  F : ARRAY[0..5931] OF REAL := [2.842882, 6.817853, 6.893808, 6.8648725, 6.890191, 6.922743, 6.92636, 6.929977, 6.9516783, 6.915509, 6.890191, 6.9733796, 6.980613, 6.890191, 6.915509, 6.919126, 6.929977, 6.9408274, 6.929977, 6.9480615, 6.991464, 7.020399, 6.9480615, 7.005932, 6.9842305, 6.9986978, 6.991464, 6.9625287, 7.005932, 7.002315, 7.0131655, 6.980613, 7.0131655, 7.0095487, 7.0131655, 6.9733796, 7.0131655, 7.0384836, 7.060185, 7.0457177, 7.096354, 7.092737, 7.0529513, 7.071036, 7.0999713, 7.0638022, 7.1180553, 7.056568, 7.1289062, 7.143374, 7.1180553, 7.1252894, 7.172309, 7.1252894, 7.1614585, 7.0891204, 7.0999713, 7.146991, 7.2229457, 7.1180553, 7.157841, 7.1903934, 7.7654805, 8.412905, 9.027778, 9.707755, 10.304543, 10.250289, 10.235822, 10.250289, 10.304543, 10.279224, 10.358796, 10.297309, 10.420283, 10.4347515, 10.373264, 10.452836, 10.456452, 10.427517, 10.463686, 10.4817705, 10.503472, 10.521557, 10.546875, 10.583044, 10.579427, 10.619213, 10.6119795, 10.644531, 10.666233, 10.734954, 10.734954, 10.698785, 10.774739, 10.78559, 10.807292, 10.778357, 10.756655, 10.821759, 10.850695, 10.807292, 10.847077, 10.904948, 10.8723955, 10.876013, 10.944734, 10.944734, 11.009838, 11.006221, 11.020689, 11.064092, 11.035156, 11.08941, 11.118345, 11.172599, 11.158131, 11.158131, 11.125579, 11.161748, 11.2630205, 11.205151, 11.29919, 11.288339, 11.219618, 11.31004, 11.306423, 11.317274, 11.349827, 11.364294, 11.378761, 11.429399, 11.447483, 11.400463, 11.454717, 11.46195, 11.490886, 11.527055, 11.548756, 11.570457, 11.624711, 11.534288, 11.682581, 11.621094, 11.599392, 11.657263, 11.747685, 11.722367, 11.76577, 11.725984, 11.71875, 11.754919, 11.801939, 11.921296, 12.008101, 12.145544, 12.286603, 12.358941, 12.398726, 12.543403, 12.641059, 12.760417, 12.814671, 12.941261, 13.057002, 13.122107, 13.208912, 13.335504, 13.440393, 13.53805, 13.599537, 13.708044, 13.791233, 13.939526, 14.022714, 14.123987, 14.210793, 14.322917, 14.391638, 14.47121, 14.579717, 14.735243, 14.728009, 14.919704, 14.999276, 15.140336, 15.223524, 15.332031, 15.4296875, 15.530961, 15.625, 15.675636, 15.838397, 15.878182, 15.921586, 16.084347, 16.24349, 16.323061, 16.44242, 16.540075, 16.543692, 16.731771, 16.818577, 16.171152, 15.386285, 14.47121, 13.729745, 12.999132, 12.890625, 12.879774, 12.97743, 12.959346, 12.959346, 13.006366, 12.999132, 13.035301, 13.006366, 13.057002, 13.075087, 13.132957, 13.132957, 13.190827, 13.198061, 13.154658, 13.266783, 13.23423, 13.28125, 13.295717, 13.299335, 13.302952, 13.317419, 13.382524, 13.349971, 13.404224, 13.483796, 13.38614, 13.505498, 13.48018, 13.530816, 13.530816, 13.581452, 13.588686, 13.6067705, 13.632089, 13.635706, 13.661024, 13.726129, 13.711661, 13.722511, 13.726129, 13.776765, 13.740596, 13.838252, 13.831018, 13.838252, 13.906974, 13.935908, 13.932292, 13.939526, 13.986546, 13.964844, 13.993779, 14.1276045, 14.019097, 14.134838, 14.134838, 14.12037, 14.138454, 14.1276045, 14.189092, 14.254195, 14.210793, 14.210793, 14.2578125, 14.290364, 14.290364, 14.348235, 14.326533, 14.395255, 14.431423, 14.420573, 14.413339, 14.478443, 14.521846, 14.507379, 14.576099, 14.514612, 14.572483, 14.58695, 14.561632, 14.699074, 14.662905, 14.69184, 14.742476, 14.767796, 14.800347, 14.78588, 14.850984, 14.803964, 16.030092, 18.514902, 21.050346, 23.488136, 25.99103, 28.47584, 30.9932, 33.449074, 35.92303, 38.465714, 40.93967, 40.990307, 37.807438, 35.337093, 32.7908, 30.35301, 27.846498, 25.343605, 22.887732, 20.330584, 17.896412, 15.379051, 13.136574, 13.111256, 13.049768, 13.111256, 13.049768, 13.0027485, 12.973814, 12.97743, 12.86169, 12.934028, 12.890625, 12.876158, 12.876158, 12.814671, 12.839989, 12.785735, 12.774884, 12.706163, 12.760417, 12.706163, 12.666377, 12.6953125, 12.644676, 12.622974, 12.597656, 12.554254, 12.590423, 12.528935, 12.503617, 12.532552, 12.510851, 12.413195, 12.420428, 12.398726, 12.402344, 12.337239, 12.351707, 12.333623, 12.261285, 12.239583, 12.257668, 12.207031, 12.203414, 12.185329, 12.163629, 12.192564, 12.141927, 12.131077, 12.047888, 12.09129, 12.040654, 12.037037, 11.982783, 12.015336, 11.961082, 11.935764, 11.92853, 11.91768, 11.856193, 11.888744, 11.867043, 11.794704, 11.801939, 11.805555, 11.762153, 11.71875, 11.700665, 11.67173, 11.697048, 11.617476, 11.584925, 11.635561, 11.599392, 11.570457, 11.555989, 11.545139, 11.516204, 11.476418, 11.498119, 11.469184, 11.46195, 11.407697, 11.342592, 11.443866, 11.349827, 11.328125, 11.281105, 11.230469, 11.306423, 11.223235, 11.201533, 11.226851, 11.129195, 11.082176, 11.111111, 11.121962, 11.078559, 11.0496235, 11.082176, 11.006221, 11.103877, 11.038774, 10.99537, 10.933883, 10.966435, 10.915798, 10.89048, 10.854311, 10.923033, 10.814526, 10.8723955, 10.767506, 10.807292, 10.796441, 10.756655, 10.713252, 10.724103, 10.655382, 10.673467, 10.6119795, 10.666233, 10.626447, 10.554109, 10.543258, 10.507089, 10.525173, 10.489005, 10.56496, 10.507089, 10.478154, 10.420283, 10.398582, 10.398582, 10.362413, 10.369647, 10.311776, 10.347945, 10.282842, 10.297309, 10.206886, 10.275608, 10.224971, 10.243055, 10.206886, 10.127315, 10.159867, 10.134548, 10.116464, 10.123698, 10.05136, 10.127315, 10.047743, 10.040509, 10.007957, 10.018807, 10.015191, 9.888599, 9.975405, 9.910301, 9.942853, 9.895833, 9.942853, 9.859664, 9.809028, 9.812645, 9.827112, 9.758391, 9.751158, 9.769242, 9.711371, 9.689671, 9.664351, 9.686053, 9.595631, 9.617332, 9.58478, 9.57393, 9.624566, 9.5703125, 9.505208, 9.4871235, 9.490741, 9.47989, 9.469039, 9.436487, 9.393085, 9.393085, 9.385851, 9.367766, 9.324364, 9.32798, 9.313513, 9.277344, 9.288195, 9.266493, 9.255642, 9.201389, 9.201389, 9.197772, 9.215857, 9.150752, 9.150752, 9.16522, 9.161603, 9.100116, 9.085649, 8.995226, 9.016927, 9.020544, 8.984375, 8.991609, 8.96629, 8.937355, 8.95544, 8.904803, 8.89757, 8.868634, 8.901186, 8.810764, 8.79268, 8.785445, 8.832465, 8.807147, 8.709491, 8.7058735, 8.723958, 8.69864, 8.676939, 8.687789, 8.637153, 8.586516, 8.669704, 8.65162, 8.311632, 7.671441, 7.060185, 6.4127603, 5.754485, 5.5266204, 5.519387, 5.541088, 5.5266204, 5.5483217, 5.46875, 5.4904513, 5.5013022, 5.4868345, 5.494068, 5.4253473, 5.4217305, 5.479601, 5.4868345, 5.396412, 5.4253473, 5.4361978, 5.428964, 5.465133, 5.4217305, 5.432581, 5.4361978, 5.443432, 5.3855615, 5.4217305, 5.4253473, 5.432581, 5.432581, 5.3855615, 5.360243, 5.4000287, 5.3493924, 5.3385415, 5.3385415, 5.331308, 5.342159, 5.342159, 5.4108796, 5.3132234, 5.360243, 5.2987556, 5.327691, 5.3023725, 5.3023725, 5.31684, 5.31684, 5.367477, 5.280671, 5.31684, 5.2842884, 5.291522, 5.255353, 5.331308, 5.2408853, 5.3132234, 5.2842884, 5.230035, 5.2842884, 5.2336516, 5.2336516, -0.014467592, 5.295139, 7.096354, 7.0493345, 7.0782695, 7.060185, 7.0240164, 7.0999713, 7.1180553, 7.0891204, 7.060185, 7.103588, 7.13614, 7.0855036, 7.1289062, 7.1252894, 7.071036, 7.1216726, 7.1903934, 7.107205, 7.1903934, 7.146991, 7.1289062, 7.146991, 7.18316, 7.1867766, 7.1650753, 7.1903934, 7.1976275, 7.18316, 7.168692, 7.2265625, 7.18316, 7.1903934, 7.212095, 7.219329, 7.208478, 7.2229457, 7.2301793, 7.1976275, 7.2554975, 7.244647, 7.2663484, 7.269965, 7.295284, 7.2229457, 7.3350697, 7.2916665, 7.284433, 7.284433, 7.2229457, 7.306134, 7.2989006, 7.280816, 7.8993053, 8.622685, 9.186921, 9.874132, 10.438368, 10.36603, 10.380498, 10.409432, 10.441985, 10.536024, 10.550492, 10.521557, 10.521557, 10.521557, 10.597511, 10.525173, 10.630064, 10.651765, 10.640914, 10.666233, 10.698785, 10.753038, 10.78559, 10.6589985, 10.789207, 10.753038, 10.814526, 10.796441, 10.810908, 10.876013, 10.865162, 10.912182, 10.908565, 10.980903, 10.912182, 10.919415, 10.98452, 10.941117, 11.017072, 11.053241, 11.031539, 11.129195, 11.107494, 11.13643, 11.121962, 11.187066, 11.201533, 11.2160015, 11.219618, 11.288339, 11.295573, 11.244936, 11.266638, 11.338976, 11.364294, 11.302807, 11.378761, 11.407697, 11.396846, 11.433015, 11.454717, 11.480035, 11.476418, 11.501736, 11.51982, 11.505353, 11.548756, 11.588542, 11.599392, 11.6066265, 11.631945, 11.610243, 11.733217, 11.71875, 11.736835, 11.700665, 11.773004, 11.834491, 11.8308735, 11.812789, 11.812789, 11.848958, 11.877893, 11.979167, 12.076823, 12.152778, 12.225116, 12.340857, 12.3878765, 12.525318, 12.641059, 12.7568, 12.894242, 12.984664, 13.0027485, 13.161892, 13.2161455, 13.3933735, 13.454861, 13.556134, 13.70081, 13.722511, 13.859954, 13.946759, 14.084202, 14.203559, 14.344618, 14.42419, 14.568866, 14.58695, 14.702691, 14.825665, 14.963108, 15.024595, 15.1222515, 15.20544, 15.328414, 15.455006, 15.534577, 15.664786, 15.769676, 15.842014, 15.983073, 16.073496, 16.210938, 16.257957, 16.37008, 16.540075, 16.597946, 16.66305, 16.847511, 16.901766, 17.035591, 17.15133, 16.88368, 15.99754, 15.133101, 14.283131, 13.415075, 12.999132, 13.053386, 13.089555, 13.118489, 13.183594, 13.125724, 13.187211, 13.165509, 13.241464, 13.208912, 13.299335, 13.313802, 13.270399, 13.299335, 13.400608, 13.364439, 13.375289, 13.43316, 13.447627, 13.451244, 13.487413, 13.494647, 13.566985, 13.516349, 13.53805, 13.610388, 13.588686, 13.661024, 13.570601, 13.751447, 13.722511, 13.7839985, 13.744213, 13.773149, 13.773149, 13.831018, 13.794849, 13.823785, 13.917824, 13.91059, 13.841869, 14.001013, 13.928675, 13.961226, 13.986546, 14.066117, 14.01548, 14.026331, 14.12037, 14.055266, 14.149305, 14.10952, 14.1746235, 14.185474, 14.26143, 14.286748, 14.27228, 14.283131, 14.337384, 14.337384, 14.398871, 14.373553, 14.416956, 14.391638, 14.496528, 14.492911, 14.492911, 14.536314, 14.550781, 14.5652485, 14.579717, 14.623119, 14.64482, 14.623119, 14.637587, 14.684607, 14.717158, 14.782263, 14.746094, 14.728009, 14.829283, 14.89077, 14.898004, 14.916088, 14.934173, 14.934173, 14.992043, 14.999276, 15.006511, 15.049913, 15.107783, 15.118634, 15.158421, 15.143952, 15.162037, 15.198206, 15.165654, 15.219908, 15.295862, 15.259693, 15.248842, 15.350116, 15.382668, 15.389901, 15.4296875, 15.400752, 15.462239, 15.47309, 15.487557, 15.563513, 17.353878, 19.889322, 22.30541, 24.833622, 27.34375, 29.78154, 32.320602, 34.776474, 37.30107, 39.803963, 42.332176, 42.306858, 38.964844, 36.433014, 33.995224, 31.488716, 29.003906, 26.450377, 24.005354, 21.538628, 18.995949, 16.53284, 14.029948, 13.237847, 13.201678, 13.183594, 13.154658, 13.154658, 13.147425, 13.132957, 13.078704, 13.042535, 13.035301, 13.006366, 13.035301, 12.973814, 12.966579, 12.854456, 12.86169, 12.850839, 12.821904, 12.792969, 12.796586, 12.771267, 12.771267, 12.771267, 12.65191, 12.630208, 12.673611, 12.662761, 12.608507, 12.637443, 12.550636, 12.554254, 12.568721, 12.474682, 12.528935, 12.39511, 12.39511, 12.3878765, 12.402344, 12.3878765, 12.311921, 12.264901, 12.282986, 12.286603, 12.246818, 12.275752, 12.217882, 12.160011, 12.170862, 12.160011, 12.145544, 12.094908, 12.062355, 12.004485, 12.029803, 11.990017, 12.000868, 11.946614, 11.932147, 11.888744, 11.859809, 11.899595, 11.874276, 11.812789, 11.841724, 11.841724, 11.769386, 11.780237, 11.762153, 11.675347, 11.642796, 11.668114, 11.67173, 11.610243, 11.581307, 11.584925, 11.537905, 11.534288, 11.555989, 11.498119, 11.411314, 11.422164, 11.436632, 11.389612, 11.34621, 11.349827, 11.378761, 11.281105, 11.302807, 11.226851, 11.252171, 11.226851, 11.201533, 11.121962, 11.165364, 11.150897, 11.114728, 11.067708, 11.056858, 11.071325, 11.024305, 11.017072, 10.970052, 10.955585, 10.959202, 10.948351, 10.883246, 10.912182, 10.865162, 10.901331, 10.796441, 10.760272, 10.763889, 10.73857, 10.720486, 10.828993, 10.73857, 10.622829, 10.677083, 10.6119795, 10.630064, 10.590278, 10.568577, 10.51794, 10.557726, 10.51794, 10.503472, 10.463686, 10.4347515, 10.449219, 10.420283, 10.380498, 10.445601, 10.304543, 10.373264, 10.286458, 10.2683735, 10.304543, 10.246673, 10.188802, 10.264757, 10.174335, 10.152633, 10.159867, 10.120081, 10.138165, 10.09838, 10.120081, 10.083912, 10.000724, 10.047743, 9.993489, 10.018807, 9.971788, 9.950087, 9.881366, 9.89945, 9.892217, 9.856048, 9.863281, 9.856048, 9.837963, 9.758391, 9.765625, 9.78371, 9.751158, 9.704138, 9.696904, 9.635417, 9.660735, 9.642651, 9.617332, 9.610099, 9.548611, 9.552228, 9.523293, 9.497974, 9.458189, 9.490741, 9.505208, 9.472656, 9.443721, 9.411169, 9.458189, 9.403935, 9.364149, 9.335214, 9.324364, 9.320746, 9.3098955, 9.237557, 9.244792, 9.201389, 9.186921, 9.212239, 9.201389, 9.132668, 9.074798, 9.060329, 9.085649, 9.035011, 9.045862, 9.060329, 8.980758, 9.00246, 8.915654, 8.904803, 8.930121, 8.861401, 8.854167, 8.839699, 8.785445, 8.828849, 8.832465, 8.774595, 8.807147, 8.691406, 8.716724, 8.687789, 8.756511, 8.666088, 8.633536, 8.622685, 8.582899, 8.553964, 8.553964, 8.557581, 8.521412, 8.525029, 8.517796, 8.496094, 8.463542, 8.420139, 8.423756, 8.39482, 8.478009, 8.391204, 8.402055, 8.340568, 8.275463, 8.293548, 8.3152485, 8.224827, 8.297164, 8.279079, 8.087384, 7.4363427, 6.7382812, 6.14511, 5.439815, 5.1576967, 5.10706, 5.0708914, 5.114294, 5.0600405, 5.1359954, 5.078125, 5.078125, 5.1215277, 5.0962095, 5.0311055, 5.0998263, 5.0455728, 5.016638, 5.0347223, 5.0311055, 5.04919, 5.013021, 5.038339, 5.038339, 5.00217, 5.027488, 4.976852, 5.00217, 5.013021, 4.9949365, 4.969618, 4.976852, 5.005787, 4.973235, 5.016638, 5.038339, 4.9949365, 4.973235, 5.013021, 4.9913197, 4.9081306, 4.9225984, 4.9334493, 4.900897, 4.864728, 4.864728, 4.9225984, 4.890046, 4.9081306, 4.8791957, 4.9153647, 4.9479165, 4.904514, 4.868345, 4.8864293, 4.8864293, 1.7216436, 2.311198, 3.0381944, 3.656684, 3.9243345, 3.8881655, 3.8809316, 3.942419, 3.9243345, 3.982205, 3.938802, 4.0256076, 3.9858217, 4.0364585, 4.0039062, 4.0364585, 4.0039062, 4.0364585, 4.0690103, 4.1377316, 4.079861, 4.0690103, 4.1341147, 4.1413484, 4.123264, 4.170284, 4.1377316, 4.1666665, 4.1304975, 4.195602, 4.181134, 4.184751, 4.260706, 4.231771, 4.2498555, 4.3113427, 4.3113427, 4.336661, 4.3185763, 4.369213, 4.3547454, 4.3402777, 4.3764467, 4.405382, 4.3909144, 4.405382, 4.448785, 4.408999, 4.4270835, 4.398148, 4.5319734, 4.5319734, 4.5572915, 4.47772, 4.5211225, 4.546441, 4.5247397, 4.5175056, 4.6006947, 4.578993, 4.571759, 4.6043115, 4.622396, 4.662182, 4.662182, 4.7200522, 4.6694155, 4.7055845, 4.763455, 4.723669, 4.7851562, 4.7417536, 4.7453704, 4.748987, 4.788773, 4.796007, 4.788773, 4.8791957, 4.835793, 4.89728, 4.8466434, 4.926215, 4.9225984, 4.8791957, 4.9153647, 4.9189816, 4.9949365, 4.9804688, 5.0094037, 4.9985533, 5.04919, 5.1576967, 5.295139, 5.403646, 5.4470487, 5.530237, 5.6278934, 5.7689524, 5.8774595, 5.9461803, 6.000434, 6.1197915, 6.1957464, 6.311487, 6.4055266, 6.4778647, 6.5827546, 6.651476, 6.752749, 6.893808, 6.9372106, 7.0457177, 7.1506076, 7.1940103, 7.316985, 7.4363427, 7.5665507, 7.5846353, 7.700376, 7.8305845, 7.8993053, 7.96441, 8.076533, 8.105469, 8.300781, 8.369502, 8.4816265, 8.532263, 8.680555, 8.7890625, 8.886719, 8.95544, 9.0494795, 9.168837, 9.248408, 9.313513, 9.469039, 9.465423, 9.6535015, 9.725839, 9.331597, 8.5286455, 7.7256947, 6.929977, 6.0800056, 5.7689524, 5.797888, 5.758102, 5.855758, 5.848524, 5.8412905, 5.83044, 5.8449073, 5.895544, 5.9534144, 5.8810763, 5.9497976, 5.9534144, 5.910012, 5.9932003, 5.9787326, 6.032986, 5.9823494, 6.0583043, 6.047454, 6.061921, 6.047454, 6.1270256, 6.0872397, 6.1306424, 6.174045, 6.1197915, 6.1306424, 6.2319155, 6.188513, 6.2029805, 6.2174478, 6.213831, 6.2355323, 6.25, 6.3440394, 6.2970195, 6.2644677, 6.358507, 6.289786, 6.3331885, 6.3187213, 6.438079, 6.3729744, 6.3729744, 6.427228, 6.4091434, 6.4453125, 6.4561634, 6.492332, 6.4850984, 6.575521, 6.514034, 6.5610533, 6.5574365, 6.5574365, 6.6840277, 6.6225405, 6.640625, 6.61169, 6.741898, 6.6948786, 6.676794, 6.7238135, 6.6731772, 6.792535, 6.7274303, 6.7853007, 6.7599826, 6.778067, 6.778067, 6.7744503, 6.8467884, 6.890191, 6.9372106, 6.850405, 6.922743, 6.9516783, 6.9335938, 6.9480615, 6.9625287, 6.980613, 6.9842305, 7.0095487, 7.027633, 7.103588, 7.0638022, 7.0746527, 7.1144385, 7.13614, 7.143374, 7.8197336, 10.300926, 12.771267, 15.295862, 17.798756, 20.283566, 22.793692, 25.296585, 27.734375, 30.197483, 32.736546, 35.232204, 37.702545, 40.227142, 40.165653, 37.08044, 34.599247, 32.08912, 29.564526, 27.155672, 24.631077, 22.128183, 19.56742, 17.126013, 14.626736, 12.163629, 9.642651, 7.1289062, 5.4108796, 5.4144964, 5.36386, 5.353009, 5.3891783, 5.3023725, 5.287905, 5.287905, 5.3240743, 5.2336516, 5.2372684, 5.280671, 5.219184, 5.219184, 5.1359954, 5.219184, 5.179398, 5.143229, 5.143229, 5.1685476, 5.074508, 5.0925927, 5.0455728, 5.0962095, 5.027488, 4.9551506, 5.0347223, 5.0094037, 5.027488, 4.9949365, 4.9804688, 4.926215, 4.9117475, 4.962384, 4.89728, 4.875579, 4.890046, 4.8466434, 4.7743053, 4.79239, 4.8213253, 4.8177085, 4.83941, 4.796007, 4.727286, 4.716435, 4.6802664, 4.7019677, 4.6875, 4.6694155, 4.647714, 4.626013, 4.651331, 4.586227, 4.636863, 4.626013, 4.539207, 4.499421, 4.560909, 4.5428243, 4.53559, 4.5319734, 4.4560184, 4.474103, 4.474103, 4.448785, 4.5211225, 4.4632525, 4.4162326, 4.3836803, 4.336661, 4.3511286, 4.296875, 4.3185763, 4.3511286, 4.3149595, 4.3041086, 4.347512, 4.2643228, 4.271557, 4.260706, 4.235388, 4.3041086, 4.1739006, 4.188368, 4.195602, 4.159433, 4.1521993, 4.119647, 4.119647, 4.108796, 4.1015625, 4.05816, 4.123264, 4.0726275, 4.083478, 3.9605036, 4.0039062, 4.007523, 4.0256076, 3.9858217, 3.8990161, 3.9568865, 3.9171007, 3.9641204, 3.9207175, 3.9026332, 3.8773148, 3.8447628, 3.8483796, 3.8447628, 3.8266783, 3.830295, 3.804977, 3.7760417, 3.7507234, 3.7000868, 3.7543402, 3.7181714, 3.7000868, 3.69647, 3.685619, 3.6892362, 3.725405, 3.6639178, 3.6385996, 3.5879629, 3.6385996, 3.5807292, 3.59158, 3.5264757, 3.5083911, 3.5228589, 3.5300925, 3.4975405, 3.5011575, 3.4324362, 3.4252026, 3.5011575, 3.4324362, 3.410735, 3.4360533, 3.3962674, 3.374566, 3.370949, 3.3673322, 3.3528645, 3.3166957, 3.378183, 3.302228, 3.2841434, 3.294994, 3.233507, 3.2732928, 3.2045717, 3.226273, 3.1864872, 3.2045717, 3.2118056, 3.1394675, 3.157552, 3.161169, 3.1358507, 3.1286168, 3.1286168, 3.0454283, 3.0635128, 3.0996816, 3.0454283, 3.049045, 3.049045, 3.023727, 3.0092592, 2.9513888, 2.9513888, 2.983941, 2.980324, 2.9296875, 2.911603, 2.8573496, 2.8645833, 2.9188368, 2.911603, 2.8175638, 2.8537326, 2.842882, 2.8320312, 2.7958622, 2.7777777, 2.8139467, 2.734375, 2.7199075, 2.7596934, 2.7162905, 2.698206, 2.7416089, 2.6945891, 2.6801214, 2.6728878, 2.6367188, 2.629485, 2.6801214, 2.6367188, 2.6150174, 2.5752316, 2.564381, 2.55353, 2.5788484, 2.5426793, 2.4920428, 2.5282118, 2.5065105, 2.5028934, 2.4775753, 2.44864, 2.4088542, 2.4233217, 2.5065105, 2.3980036, 2.445023, 2.3582175, 2.4233217, 2.3618345, 2.376302, 2.3654513, 2.2858796, 2.3184316, 2.23886, 2.3365161, 2.275029, 2.2605612, 2.1918402, 2.2280092, 1.634838, 0.9765625, 0.30020255, 3.4432871, 5.0455728, 5.0998263, 5.10706, 5.0853586, 5.1613135, 5.117911, 5.128762, 5.0925927, 5.143229, 5.0600405, 5.0708914, 5.1649303, 5.128762, 5.114294, 5.103443, 5.1576967, 5.183015, 5.117911, 5.1576967, 5.179398, 5.1649303, 5.0708914, 5.1251445, 5.215567, 5.179398, 5.2119503, 5.1721644, 5.204716, 5.150463, 5.204716, 5.179398, 5.190249, 5.1974826, 5.2445025, 5.2408853, 5.1757812, 5.251736, 5.280671, 5.2445025, 5.255353, 5.2842884, 5.2408853, 5.280671, 5.2445025, 5.2336516, 5.2987556, 5.230035, 5.2698207, 5.31684, 5.3783274, 5.3385415, 5.2987556, 5.287905, 5.3132234, 5.2770543, 5.3747106, 5.3132234, 5.4000287, 5.353009, 5.3096066, 5.6315103, 6.3368053, 6.969763, 7.60272, 8.282697, 8.427373, 8.405671, 8.445457, 8.456307, 8.423756, 8.510561, 8.539496, 8.564815, 8.496094, 8.59375, 8.600984, 8.619068, 8.557581, 8.691406, 8.669704, 8.691406, 8.738426, 8.637153, 8.763744, 8.781829, 8.796296, 8.785445, 8.80353, 8.843316, 8.854167, 8.875868, 8.843316, 8.908421, 8.937355, 8.9192705, 9.006077, 8.959057, 8.998842, 8.973524, 9.016927, 9.031395, 9.031395, 8.998842, 9.085649, 9.063947, 9.154369, 9.186921, 9.161603, 9.273726, 9.201389, 9.226707, 9.233941, 9.248408, 9.248408, 9.338831, 9.338831, 9.349682, 9.302662, 9.364149, 9.447338, 9.367766, 9.454572, 9.385851, 9.42202, 9.476274, 9.490741, 9.505208, 9.505208, 9.602864, 9.555845, 9.544994, 9.588397, 9.628182, 9.664351, 9.628182, 9.660735, 9.682436, 9.729456, 9.707755, 9.73669, 9.740307, 9.823495, 9.805411, 9.798177, 9.823495, 9.866899, 9.881366, 9.85243, 9.975405, 10.007957, 9.95732, 10.029658, 10.185185, 10.206886, 10.315393, 10.467303, 10.554109, 10.691551, 10.756655, 10.789207, 10.966435, 11.067708, 11.161748, 11.205151, 11.338976, 11.472801, 11.555989, 11.603009, 11.715133, 11.794704, 11.924913, 12.040654, 12.131077, 12.203414, 12.355324, 12.384259, 12.507234, 12.60489, 12.648293, 12.800202, 12.9557295, 13.042535, 13.078704, 13.165509, 13.32827, 13.404224, 13.527199, 13.58507, 13.726129, 13.820168, 13.968461, 13.990162, 14.134838, 14.21441, 14.279514, 14.362702, 14.532697, 14.619502, 14.7316265, 14.840133, 14.923322, 14.623119, 13.798467, 12.9557295, 12.160011, 11.382379, 11.020689, 11.053241, 11.121962, 11.107494, 11.143663, 11.121962, 11.150897, 11.14728, 11.219618, 11.190682, 11.183449, 11.223235, 11.302807, 11.295573, 11.255787, 11.364294, 11.317274, 11.375145, 11.3932295, 11.418548, 11.4402485, 11.469184, 11.436632, 11.494502, 11.494502, 11.588542, 11.555989, 11.559607, 11.603009, 11.617476, 11.617476, 11.704283, 11.693432, 11.678964, 11.715133, 11.744068, 11.773004, 11.758536, 11.816406, 11.809173, 11.848958, 11.910445, 11.950232, 11.874276, 11.932147, 11.924913, 11.968316, 11.979167, 12.004485, 12.037037, 12.000868, 12.123842, 12.105758, 12.181713, 12.141927, 12.203414, 12.13831, 12.203414, 12.239583, 12.250434, 12.2432, 12.29022, 12.326389, 12.366175, 12.362557, 12.358941, 12.3878765, 12.3878765, 12.424046, 12.405961, 12.485533, 12.528935, 12.528935, 12.528935, 12.54702, 12.554254, 12.615741, 12.619358, 12.626592, 12.662761, 12.6953125, 12.764033, 12.811053, 12.724248, 12.760417, 12.80382, 12.843605, 12.836371, 12.850839, 12.90871, 12.941261, 13.292101, 15.704572, 18.17853, 20.706741, 23.1807, 25.672743, 28.121384, 30.671297, 33.15249, 35.633682, 38.151043, 40.588833, 40.559895, 37.492767, 34.964554, 32.508682, 30.016638, 27.50651, 25.043404, 22.518808, 20.070168, 17.520254, 15.089699, 12.579572, 11.237702, 11.161748, 11.2160015, 11.114728, 11.100261, 11.121962, 11.096643, 11.085793, 11.031539, 11.024305, 11.056858, 10.951967, 11.020689, 10.944734, 10.912182, 10.901331, 10.87963, 10.8253765, 10.803675, 10.789207, 10.73857, 10.745805, 10.781974, 10.706018, 10.724103, 10.593895, 10.673467, 10.6807, 10.572193, 10.554109, 10.579427, 10.503472, 10.521557, 10.52879, 10.463686, 10.445601, 10.46007, 10.532408, 10.420283, 10.35518, 10.322627, 10.326244, 10.3515625, 10.286458, 10.250289, 10.243055, 10.228588, 10.2213545, 10.181568, 10.206886, 10.192419, 10.083912, 10.112847, 10.083912, 10.054976, 10.047743, 10.007957, 10.007957, 9.964555, 9.982639, 9.986256, 9.924768, 9.89945, 9.892217, 9.848814, 9.837963, 9.884983, 9.801794, 9.780092, 9.780092, 9.754774, 9.725839, 9.725839, 9.711371, 9.693287, 9.6535015, 9.617332, 9.628182, 9.599248, 9.566695, 9.610099, 9.57393, 9.508825, 9.4871235, 9.443721, 9.414786, 9.43287, 9.382234, 9.382234, 9.360533, 9.324364, 9.338831, 9.306279, 9.378617, 9.244792, 9.215857, 9.2628765, 9.291811, 9.186921, 9.183305, 9.190538, 9.194155, 9.147136, 9.067564, 9.035011, 9.009693, 9.103733, 8.991609, 9.009693, 9.009693, 8.991609, 9.027778, 8.933739, 8.8722515, 8.933739, 8.865017, 8.875868, 8.843316, 8.7890625, 8.843316, 8.74566, 8.713108, 8.767361, 8.7058735, 8.687789, 8.673322, 8.7058735, 8.600984, 8.597367, 8.604601, 8.600984, 8.575665, 8.532263, 8.532263, 8.521412, 8.553964, 8.5286455, 8.478009, 8.4816265, 8.470776, 8.409288, 8.351418, 8.308015, 8.362268, 8.3152485, 8.3152485, 8.297164, 8.293548, 8.213976, 8.206742, 8.199508, 8.224827, 8.192274, 8.17419, 8.18504, 8.134404, 8.101851, 8.065682, 8.080151, 8.065682, 8.065682, 8.025897, 7.9716434, 8.036748, 7.9318576, 7.939091, 7.949942, 7.913773, 7.9029226, 7.8703704, 7.884838, 7.8956885, 7.837818, 7.8052664, 7.747396, 7.7582464, 7.7256947, 7.7546296, 7.703993, 7.6931424, 7.7293115, 7.6678243, 7.6171875, 7.5882525, 7.6497397, 7.5810184, 7.573785, 7.5810184, 7.530382, 7.5520835, 7.5050635, 7.486979, 7.472512, 7.5014467, 7.396557, 7.382089, 7.458044, 7.360388, 7.3423033, 7.349537, 7.309751, 7.3025174, 7.248264, 7.306134, 7.269965, 7.2265625, 7.1903934, 7.157841, 7.2012444, 7.139757, 7.168692, 7.1108217, 7.081887, 7.0746527, 7.0999713, 7.0457177, 7.1759257, 7.027633, 7.03125, 6.9878473, 6.9733796, 7.0131655, 6.929977, 6.8757234, 6.8974247, 6.857639, 6.8467884, 6.8865743, 6.8106194, 6.7599826, 6.792535, 6.814236, 6.792535, 6.2970195, 5.6351275, 4.875579, 4.257089, 3.6639178, 3.7073207, 3.69647, 3.6385996, 3.692853, 3.685619, 3.660301, 3.6639178, 3.6385996, 3.656684, 3.7181714, 3.685619, 3.6422164, 3.6277487, 3.620515, 3.6458333, 3.6385996, 3.5951967, 3.584346, 3.6313658, 3.5988138, 3.5879629, 3.5807292, 3.5879629, 3.5554109, 3.5879629, 3.59158, 3.551794, 3.5300925, 3.6060474, 3.5554109, 3.5300925, 3.5409434, 3.5264757, 3.5047743, 3.5192418, 3.5083911, 3.5373263, 3.5626447, 3.5011575, 3.5409434, 3.4866898, 3.5662615, 3.5120082, 3.5047743, 3.5192418, 3.4903066, 3.5228589, 3.4866898, 3.4505208, 3.4722223, 3.4649885, 3.446904, 3.4577546, 3.3528645, 3.4939237, 3.4866898, 3.4179688, 3.4215856, 3.4252026, 3.378183, 1.8916377, 4.615162, 4.626013, 4.5645256, 4.6187787, 4.6187787, 4.560909, 4.662182, 4.6296296, 4.6187787, 4.615162, 4.5645256, 4.622396, 4.6079283, 4.658565, 4.683883, 4.622396, 4.6043115, 4.691117, 4.6875, 4.676649, 4.647714, 4.6440973, 4.651331, 4.691117, 4.5898438, 4.6043115, 4.6730323, 4.723669, 4.6332464, 4.6730323, 4.7019677, 4.727286, 4.698351, 4.7019677, 4.6875, 4.6802664, 4.6730323, 4.6802664, 4.716435, 4.6947336, 4.6549478, 4.727286, 4.7345195, 4.738137, 4.727286, 4.788773, 4.7815394, 4.788773, 4.7670717, 4.7706885, 4.799624, 4.738137, 4.738137, 4.8177085, 4.763455, 4.8574944, 4.7815394, 4.7670717, 4.796007, 4.803241, 4.9479165, 5.5917244, 6.2934027, 6.919126, 7.526765, 7.8956885, 7.8920717, 7.8920717, 7.939091, 7.9029226, 7.960793, 7.960793, 7.960793, 7.9788775, 7.96441, 7.9463253, 8.036748, 8.018663, 8.087384, 8.065682, 8.105469, 8.141638, 8.188658, 8.145255, 8.181423, 8.192274, 8.17419, 8.275463, 8.206742, 8.199508, 8.308015, 8.257379, 8.311632, 8.326099, 8.33695, 8.322483, 8.33695, 8.3152485, 8.412905, 8.380353, 8.344184, 8.463542, 8.412905, 8.467158, 8.459925, 8.525029, 8.496094, 8.499711, 8.568432, 8.499711, 8.575665, 8.564815, 8.619068, 8.626302, 8.684173, 8.629919, 8.684173, 8.69864, 8.662471, 8.713108, 8.716724, 8.785445, 8.774595, 8.785445, 8.7890625, 8.79268, 8.846932, 8.825232, 8.904803, 8.890336, 8.930121, 8.987992, 8.973524, 8.944589, 8.933739, 9.07118, 9.01331, 9.038629, 9.020544, 9.056713, 9.07118, 9.038629, 9.125434, 9.1182, 9.103733, 9.190538, 9.139901, 9.215857, 9.244792, 9.226707, 9.284577, 9.302662, 9.400318, 9.519676, 9.602864, 9.696904, 9.801794, 9.870515, 9.94647, 10.058594, 10.174335, 10.275608, 10.380498, 10.456452, 10.568577, 10.698785, 10.745805, 10.836226, 10.944734, 11.078559, 11.085793, 11.248553, 11.367911, 11.458333, 11.530671, 11.621094, 11.700665, 11.841724, 11.92853, 12.029803, 12.152778, 12.207031, 12.344474, 12.377026, 12.518085, 12.637443, 12.713397, 12.811053, 12.883391, 13.064236, 13.089555, 13.22338, 13.292101, 13.436776, 13.527199, 13.610388, 13.718895, 13.820168, 13.932292, 14.001013, 14.073351, 13.943142, 13.136574, 12.380642, 11.563224, 10.662616, 10.199653, 10.206886, 10.275608, 10.264757, 10.257524, 10.271991, 10.282842, 10.322627, 10.402199, 10.3515625, 10.36603, 10.423901, 10.470921, 10.489005, 10.478154, 10.536024, 10.525173, 10.521557, 10.539641, 10.568577, 10.622829, 10.604745, 10.640914, 10.63368, 10.615596, 10.6589985, 10.698785, 10.767506, 10.687934, 10.724103, 10.78559, 10.807292, 10.854311, 10.756655, 10.821759, 10.774739, 10.876013, 10.857928, 10.894097, 10.857928, 10.926649, 10.930266, 10.988136, 11.035156, 11.046007, 11.038774, 11.017072, 11.096643, 11.118345, 11.085793, 11.143663, 11.201533, 11.1943, 11.201533, 11.176215, 11.230469, 11.205151, 11.342592, 11.291956, 11.31004, 11.313658, 11.313658, 11.331742, 11.41493, 11.443866, 11.407697, 11.46195, 11.447483, 11.490886, 11.51982, 11.541522, 11.545139, 11.501736, 11.628327, 11.621094, 11.628327, 11.639178, 11.624711, 11.646412, 11.682581, 11.729601, 11.71875, 11.791088, 11.794704, 11.856193, 11.834491, 11.780237, 11.845342, 11.852575, 11.859809, 11.932147, 12.084057, 14.369936, 16.880064, 19.382957, 21.849682, 24.374277, 26.837385, 29.394531, 31.807003, 34.324364, 36.816406, 39.304832, 41.82581, 41.822193, 38.697193, 36.23047, 33.716724, 31.210215, 28.68562, 26.182726, 23.672598, 21.216724, 18.75, 16.26519, 13.75868, 11.2160015, 10.21412, 10.170717, 10.199653, 10.116464, 10.058594, 10.112847, 10.073061, 10.10923, 10.080296, 9.993489, 10.015191, 10.040509, 9.968171, 9.928386, 9.924768, 9.982639, 9.942853, 9.859664, 9.870515, 9.845197, 9.845197, 9.834346, 9.85243, 9.686053, 9.765625, 9.725839, 9.73669, 9.718605, 9.7005205, 9.671586, 9.628182, 9.613715, 9.599248, 9.508825, 9.519676, 9.508825, 9.47989, 9.530526, 9.505208, 9.4401045, 9.461805, 9.458189, 9.396702, 9.360533, 9.389467, 9.295428, 9.331597, 9.306279, 9.284577, 9.313513, 9.233941, 9.295428, 9.230324, 9.226707, 9.215857, 9.136285, 9.129051, 9.0964985, 9.1182, 9.0964985, 9.056713, 9.085649, 9.042245, 9.016927, 8.998842, 9.006077, 8.959057, 8.995226, 8.933739, 8.886719, 8.868634, 8.868634, 8.886719, 8.861401, 8.825232, 8.846932, 8.723958, 8.7890625, 8.74566, 8.716724, 8.676939, 8.64077, 8.695024, 8.65162, 8.637153, 8.648004, 8.64077, 8.615452, 8.586516, 8.568432, 8.539496, 8.539496, 8.470776, 8.532263, 8.423756, 8.430989, 8.44184, 8.365886, 8.485243, 8.344184, 8.373119, 8.304399, 8.355035, 8.3152485, 8.300781, 8.246528, 8.297164, 8.257379, 8.235677, 8.206742, 8.199508, 8.177807, 8.159722, 8.152489, 8.065682, 8.148871, 8.083767, 8.065682, 8.051215, 8.047599, 8.029514, 8.01143, 7.9824944, 7.9571757, 7.9427085, 7.921007, 7.924624, 7.888455, 7.8956885, 7.8450522, 7.816117, 7.8305845, 7.873987, 7.7944155, 7.7980323, 7.675058, 7.751013, 7.736545, 7.675058, 7.6569734, 7.7329283, 7.664207, 7.6822915, 7.624421, 7.624421, 7.599103, 7.5810184, 7.5774016, 7.533999, 7.494213, 7.548466, 7.4652777, 7.530382, 7.4905963, 7.3893228, 7.411024, 7.3676214, 7.458044, 7.411024, 7.3350697, 7.3314524, 7.313368, 7.309751, 7.3025174, 7.2663484, 7.284433, 7.2374134, 7.233796, 7.244647, 7.219329, 7.132523, 7.143374, 7.143374, 7.096354, 7.0746527, 7.1289062, 7.0638022, 7.1252894, 7.0529513, 7.0638022, 7.027633, 6.9444447, 7.0638022, 6.9769964, 6.9408274, 6.966146, 6.9625287, 6.893808, 6.9625287, 6.890191, 6.890191, 6.8721066, 6.8359375, 6.8033853, 6.7997684, 6.745515, 6.749132, 6.781684, 6.702112, 6.7853007, 6.7382812, 6.7093463, 6.6731772, 6.629774, 6.6478586, 6.589988, 6.6080728, 6.6623263, 6.604456, 6.5502024, 6.5502024, 6.528501, 6.4742475, 6.503183, 6.463397, 6.4561634, 6.430845, 6.4199944, 6.4344616, 6.488715, 6.3946757, 6.391059, 6.311487, 6.351273, 6.3187213, 6.351273, 6.3078704, 6.275318, 6.2825522, 6.300637, 6.2355323, 6.25, 6.1957464, 5.5157695, 4.9189816, 4.235388, 3.6639178, 3.1394675, 3.125, 3.125, 3.092448, 3.0996816, 3.1141493, 3.1141493, 3.1213832, 3.0743635, 3.1032987, 3.092448, 3.1141493, 3.0996816, 3.1286168, 3.0381944, 3.1177661, 3.1539352, 3.0996816, 3.0635128, 3.0779803, 3.1032987, 3.0743635, 3.0309606, 3.02011, 3.0960648, 3.0635128, 3.092448, 3.0418112, 3.0526621, 3.0454283, 3.0707464, 3.0309606, 3.0345776, 3.0273438, 3.0128763, 3.0671296, 3.0020254, 3.0418112, 3.0526621, 2.9911747, 2.983941, 3.016493, 3.0598958, 3.0598958, 3.0418112, 2.9947917, 2.9911747, 3.0020254, 3.023727, 2.9911747, 2.9947917, 3.0056424, 2.9947917, 2.9767072, 2.947772, 2.9694734, 2.9694734, 2.947772, 2.9730902, 3.023727, 0.003616898, 3.8917825, 7.8667536, 10.387732, 10.405816, 10.4347515, 10.358796, 10.4347515, 10.423901, 10.423901, 10.405816, 10.391349, 10.441985, 10.423901, 10.427517, 10.445601, 10.46007, 10.463686, 10.507089, 10.4347515, 10.427517, 10.496239, 10.456452, 10.478154, 10.463686, 10.496239, 10.496239, 10.4817705, 10.416667, 10.499855, 10.51794, 10.525173, 10.532408, 10.489005, 10.507089, 10.532408, 10.496239, 10.52879, 10.590278, 10.507089, 10.550492, 10.543258, 10.561342, 10.604745, 10.590278, 10.57581, 10.601129, 10.554109, 10.543258, 10.57581, 10.604745, 10.666233, 10.640914, 10.604745, 10.6119795, 10.622829, 10.6119795, 10.63368, 10.637298, 10.669849, 10.6589985, 10.626447, 10.6807, 10.912182, 11.490886, 12.087673, 12.807436, 13.472945, 13.718895, 13.733362, 13.75868, 13.827401, 13.834636, 13.878038, 13.8671875, 13.906974, 13.86357, 13.896123, 13.928675, 13.982928, 13.964844, 14.00463, 13.939526, 14.037182, 14.033565, 14.102286, 14.1276045, 14.080585, 14.1276045, 14.102286, 14.171007, 14.156539, 14.1746235, 14.210793, 14.221643, 14.265046, 14.239728, 14.268663, 14.279514, 14.333767, 14.297599, 14.312066, 14.355469, 14.362702, 14.406105, 14.402489, 14.409722, 14.514612, 14.48206, 14.500145, 14.510995, 14.456742, 14.525463, 14.561632, 14.63397, 14.58695, 14.615886, 14.63397, 14.688224, 14.655671, 14.670139, 14.713542, 14.709925, 14.775029, 14.782263, 14.800347, 14.811198, 14.847367, 14.9088545, 14.854601, 14.869068, 14.90162, 14.934173, 14.923322, 14.959491, 14.945024, 15.002893, 15.028212, 15.05353, 15.0390625, 15.071614, 15.060764, 15.075232, 15.143952, 15.140336, 15.165654, 15.172888, 15.194589, 15.212673, 15.237992, 15.230758, 15.274161, 15.292245, 15.259693, 15.436921, 15.47309, 15.56713, 15.704572, 15.809462, 15.925202, 15.99754, 16.040943, 16.229021, 16.29051, 16.413485, 16.45327, 16.594328, 16.735388, 16.771557, 16.945168, 16.974104, 17.086227, 17.126013, 17.256222, 17.386429, 17.520254, 17.563658, 17.690248, 17.82769, 17.914497, 17.939816, 18.051939, 18.171297, 18.254484, 18.381077, 18.525753, 18.612558, 18.663195, 18.757235, 18.898293, 18.981482, 19.089989, 19.245516, 19.288918, 19.433594, 19.560184, 19.599972, 19.62529, 19.806135, 19.896557, 19.979746, 20.120804, 20.225695, 20.330584, 20.272715, 19.480614, 18.565538, 17.856627, 17.006655, 16.485823, 16.44242, 16.550926, 16.456886, 16.540075, 16.56901, 16.554543, 16.608797, 16.597946, 16.659433, 16.71007, 16.724537, 16.735388, 16.677517, 16.728153, 16.735388, 16.861979, 16.796875, 16.83666, 16.847511, 16.854746, 16.912615, 16.876448, 16.959635, 17.006655, 16.934317, 16.988571, 16.988571, 17.01389, 17.089844, 17.158566, 17.078993, 17.158566, 17.122396, 17.205584, 17.227285, 17.24537, 17.216434, 17.238136, 17.31409, 17.30324, 17.364729, 17.346643, 17.433449, 17.4443, 17.415365, 17.386429, 17.404514, 17.45515, 17.509403, 17.534721, 17.574509, 17.574509, 17.545572, 17.603443, 17.635996, 17.668547, 17.730034, 17.733652, 17.730034, 17.766203, 17.831308, 17.798756, 17.849392, 17.824074, 17.914497, 17.892796, 17.939816, 17.943432, 18.00492, 18.019386, 18.041088, 18.055555, 18.023003, 18.091724, 18.149595, 18.124277, 18.185764, 18.214699, 18.17853, 18.2364, 18.258102, 18.27257, 18.315971, 18.315971, 18.381077, 18.359375, 18.370226, 18.471498, 18.48235, 18.467882, 18.4932, 20.554832, 23.021557, 25.56062, 27.987558, 30.50492, 33.062065, 35.467304, 37.94126, 40.46224, 40.505642, 36.4511, 32.461662, 29.644096, 27.083334, 24.660011, 22.063078, 19.632523, 17.111546, 14.594184, 12.149161, 9.8307295, 9.42202, 9.497974, 9.436487, 9.360533, 9.367766, 9.302662, 9.299046, 9.2628765, 9.324364, 9.230324, 9.2628765, 9.201389, 9.248408, 9.161603, 9.139901, 9.129051, 9.129051, 9.053096, 9.082031, 9.038629, 9.01331, 8.987992, 8.95544, 8.940972, 8.940972, 8.9192705, 8.904803, 8.901186, 8.915654, 8.828849, 8.832465, 8.810764, 8.79268, 8.738426, 8.752893, 8.749276, 8.65162, 8.669704, 8.65162, 8.626302, 8.586516, 8.633536, 8.575665, 8.586516, 8.5286455, 8.470776, 8.434607, 8.430989, 8.478009, 8.409288, 8.365886, 8.33695, 8.409288, 8.333333, 8.344184, 8.347801, 8.318866, 8.322483, 8.308015, 8.192274, 8.250145, 8.206742, 8.192274, 8.163339, 8.058449, 8.105469, 8.112702, 8.047599, 8.029514, 8.080151, 8.015046, 8.0078125, 7.91739, 8.015046, 7.9318576, 7.8956885, 7.8993053, 7.8667536, 7.928241, 7.837818, 7.9065394, 7.7690973, 7.837818, 7.7907987, 7.7437787, 7.7437787, 7.740162, 7.664207, 7.7220774, 7.635272, 7.609954, 7.6063366, 7.6280384, 7.573785, 7.5665507, 7.5159144, 7.5014467, 7.4544272, 7.5050635, 7.4761286, 7.425492, 7.4399595, 7.39294, 7.411024, 7.385706, 7.3350697, 7.3350697, 7.3386865, 7.273582, 7.284433, 7.2663484, 7.2301793, 7.2157116, 7.1976275, 7.157841, 7.1940103, 7.1867766, 7.139757, 7.1144385, 7.096354, 7.081887, 7.0638022, 7.034867, 7.060185, 6.9842305, 6.854022, 6.980613, 6.9408274, 6.929977, 6.904659, 6.9118924, 6.82147, 6.828704, 6.817853, 6.778067, 6.7961516, 6.7310476, 6.7853007, 6.778067, 6.702112, 6.665943, 6.680411, 6.629774, 6.579138, 6.6225405, 6.6550927, 6.5863714, 6.640625, 6.5502024, 6.5610533, 6.514034, 6.467014, 6.4814816, 6.4959493, 6.45978, 6.430845, 6.391059, 6.35489, 6.391059, 6.358507, 6.362124, 6.35489, 6.35489, 6.289786, 6.25, 6.1921296, 6.239149, 6.221065, 6.1921296, 6.1704283, 6.1306424, 6.1631947, 6.1306424, 6.112558, 6.141493, 6.069155, 6.0149016, 6.0257525, 6.0149016, 5.9136286, 5.996817, 5.964265, 5.920862, 5.964265, 5.862992, 5.9136286, 5.870226, 5.8521414, 5.834057, 5.8521414, 5.808738, 5.794271, 5.797888, 5.7725697, 5.7038484, 5.721933, 5.6893806, 5.6532116, 5.721933, 5.67853, 5.6387444, 5.6025753, 5.5664062, 5.5627894, 5.5013022, 5.5483217, 5.4832177, 5.497685, 5.497685, 5.4615164, 5.479601, 5.443432, 5.4361978, 5.392795, 5.3819447, 5.3710938, 5.327691, 5.255353, 5.3132234, 5.2408853, 5.186632, 5.291522, 5.2481194, 5.2372684, 5.2372684, 5.2010994, 5.1974826, 5.1721644, 5.1757812, 5.15408, 5.15408, 5.0962095, 4.9153647, 4.2426214, 3.584346, 2.983941, 2.3039641, 2.0182292, 1.9675926, 1.9929109, 2.0073786, 2.0146122, 1.9748263, 1.9856771, 1.9024885, 1.9712095, 1.8952546, 1.9675926, 1.9748263, 1.9241898, 1.9567419, 1.9458913, 1.9422743, 1.9748263, 1.8735533, 1.9024885, 1.9205729, 1.9241898, 1.9133391, 1.880787, 1.9350405, 1.9567419, 1.8590857, 1.9024885, 1.8880209, 1.8373842, 1.8590857, 1.884404, 1.8699363, 1.8265336, 1.8229166, 1.812066, 1.8554688, 1.8554688, 1.848235, 1.848235, 1.8590857, 1.8265336, 1.775897, 1.8446181, 1.8192998, 1.7903646, 1.8301505, 1.8554688, 1.7903646, 1.739728, 1.8012153, 1.7614294, 1.808449, 1.775897, 1.7469618, 1.7505788, 1.8012153, 1.7650462, 1.7722801, 1.7433449, 1.775897, 2.665654, 6.741898, 6.904659, 6.915509, 6.980613, 6.9625287, 6.8612556, 6.958912, 6.904659, 6.8721066, 6.922743, 6.9372106, 6.929977, 6.955295, 6.9372106, 6.87934, 6.904659, 6.9625287, 6.966146, 6.922743, 6.9625287, 6.92636, 6.958912, 7.0167823, 6.966146, 7.071036, 6.958912, 7.002315, 6.969763, 6.9769964, 6.9842305, 7.0131655, 7.005932, 7.020399, 7.0999713, 7.067419, 7.0384836, 7.0240164, 7.0167823, 7.0384836, 7.060185, 7.0782695, 7.0999713, 7.071036, 7.139757, 7.0891204, 7.0384836, 7.081887, 7.103588, 7.1614585, 7.1216726, 7.1180553, 7.092737, 7.157841, 7.1542244, 7.13614, 7.1614585, 7.107205, 7.18316, 7.146991, 7.2012444, 7.1940103, 7.1903934, 7.107205, 7.2012444, 7.1506076, 7.18316, 7.179543, 7.1903934, 7.1903934, 7.233796, 7.1940103, 7.2012444, 7.2157116, 7.2012444, 7.204861, 7.2518806, 7.269965, 7.2157116, 7.2229457, 7.244647, 7.2916665, 7.24103, 7.2916665, 7.295284, 7.295284, 7.2627316, 7.2518806, 7.3025174, 7.3025174, 7.306134, 7.24103, 7.2916665, 7.313368, 7.418258, 7.3242188, 7.4001737, 7.284433, 7.349537, 7.3386865, 7.3278356, 7.3784723, 7.313368, 7.425492, 7.3748555, 7.3784723, 7.4074073, 7.3640046, 7.418258, 7.4291086, 7.3640046, 7.4001737, 7.421875, 7.3784723, 7.4399595, 7.45081, 7.4037905, 7.4291086, 7.4001737, 7.4652777, 7.4761286, 7.458044, 7.472512, 7.4761286, 7.5014467, 7.4797454, 7.5014467, 7.4363427, 7.4761286, 7.5014467, 7.5159144, 7.5195312, 7.486979, 7.526765, 7.5448494, 7.533999, 7.5448494, 7.570168, 7.5520835, 7.548466, 7.548466, 7.5557003, 7.562934, 7.559317, 7.5810184, 7.60272, 7.526765, 7.5557003, 7.595486, 7.5882525, 7.6533566, 7.6171875, 7.6171875, 7.6425056, 7.6497397, 7.6280384, 7.6497397, 7.6533566, 7.6822915, 7.6533566, 7.703993, 7.696759, 7.70761, 7.6822915, 7.675058, 7.696759, 7.7582464, 7.7220774, 7.6931424, 7.7220774, 7.7329283, 7.7582464, 7.7546296, 7.7220774, 7.7293115, 7.7582464, 7.7293115, 7.761863, 7.7437787, 7.7256947, 7.7582464, 7.7980323, 7.7944155, 7.772714, 7.8595195, 7.837818, 7.8305845, 7.7980323, 7.877604, 7.837818, 7.8812213, 7.9354744, 7.877604, 7.921007, 7.8812213, 7.9029226, 7.949942, 7.8956885, 7.888455, 7.921007, 7.873987, 7.913773, 7.8920717, 7.924624, 7.939091, 7.9354744, 7.939091, 7.9571757, 7.949942, 7.9716434, 7.96441, 7.9824944, 8.02228, 7.993345, 8.047599, 7.989728, 7.986111, 8.058449, 8.015046, 8.087384, 7.9788775, 8.029514, 8.029514, 8.015046, 8.051215, 8.000579, 8.065682, 8.036748, 8.101851, 8.130787, 8.0910015, 8.098235, 8.087384, 8.109086, 8.134404, 8.072917, 8.130787, 8.152489, 8.159722, 8.159722, 8.141638, 8.181423, 8.152489, 8.134404, 8.18504, 8.156105, 8.253761, 8.210359, 8.206742, 8.286314, 8.250145, 8.264612, 8.239294, 8.250145, 8.264612, 8.257379, 8.28993, 8.28993, 8.260995, 8.2682295, 8.326099, 8.3152485, 8.39482, 8.322483, 8.293548, 8.297164, 8.308015, 8.344184, 8.369502, 8.333333, 8.412905, 8.39482, 8.402055, 8.402055, 8.467158, 8.412905, 8.412905, 8.420139, 8.423756, 8.463542, 8.456307, 8.449074, 8.391204, 8.53588, 8.459925, 8.496094, 8.48886, 8.430989, 8.532263, 8.510561, 8.474392, 8.53588, 8.525029, 8.582899, 8.525029, 8.532263, 8.550347, 8.770978, 11.060474, 13.581452, 16.04456, 18.518518, 21.097366, 23.53154, 26.016348, 28.468605, 31.011284, 33.52141, 35.991753, 38.43316, 40.91797, 40.99754, 37.7785, 35.380497, 32.816116, 30.349392, 27.81033, 25.347221, 22.858797, 20.413773, 17.86386, 15.350116, 12.91956, 10.376881, 7.96441, 6.8250866, 6.8612556, 6.8106194, 6.8359375, 6.8395543, 6.8106194, 6.792535, 6.8106194, 6.7744503, 6.7853007, 6.792535, 6.756366, 6.7744503, 6.7274303, 6.7382812, 6.756366, 6.767216, 6.749132, 6.6876445, 6.7635994, 6.7708335, 6.7093463, 6.702112, 6.741898, 6.691262, 6.640625, 6.6948786, 6.6333914, 6.640625, 6.604456, 6.651476, 6.640625, 6.6478586, 6.600839, 6.5936055, 6.6080728, 6.5863714, 6.5863714, 6.6080728, 6.6225405, 6.6189237, 6.579138, 6.615307, 6.6080728, 6.5610533, 6.6225405, 6.528501, 6.5502024, 6.524884, 6.492332, 6.528501, 6.5104165, 6.532118, 6.4453125, 6.488715, 6.4489293, 6.488715, 6.4778647, 6.4706306, 6.463397, 6.40191, 6.4344616, 6.4453125, 6.4416957, 6.4489293, 6.387442, 6.4091434, 6.423611, 6.40191, 6.427228, 6.427228, 6.3946757, 6.376591, 6.45978, 6.3729744, 6.351273, 6.2970195, 6.3838253, 6.358507, 6.325955, 6.3331885, 6.289786, 6.322338, 6.3693576, 6.3295717, 6.2934027, 6.2825522, 6.3042536, 6.325955, 6.184896, 6.260851, 6.2644677, 6.2970195, 6.2174478, 6.2319155, 6.1921296, 6.25, 6.2427664, 6.2029805, 6.210214, 6.199363, 6.239149, 6.184896, 6.213831, 6.1957464, 6.1631947, 6.239149, 6.1559606, 6.1559606, 6.2065973, 6.0872397, 6.1668115, 6.174045, 6.148727, 6.101707, 6.188513, 6.1595774, 6.069155, 6.148727, 6.112558, 6.0944734, 6.0836225, 6.047454, 6.0836225, 6.061921, 6.09809, 6.0872397, 6.061921, 6.1197915, 6.0655384, 6.061921, 6.0185184, 6.0944734, 6.047454, 6.032986, 6.04022, 6.007668, 5.985966, 6.007668, 6.0221353, 5.985966, 5.960648, 5.996817, 5.964265, 5.975116, 6.0293694, 6.0221353, 5.9497976, 5.9570312, 5.964265, 6.0040507, 5.931713, 5.9136286, 5.9497976, 5.924479, 5.9425635, 5.9280963, 5.9136286, 5.8810763, 5.870226, 5.8810763, 5.8412905, 5.9280963, 5.8449073, 5.8449073, 5.8774595, 5.8376737, 5.823206, 5.8810763, 5.855758, 5.855758, 5.797888, 5.8123555, 5.8738427, 5.7761865, 5.7725697, 5.8376737, 5.78342, 5.743634, 5.808738, 5.732784, 5.8051214, 5.7761865, 5.747251, 5.78342, 5.743634, 5.8015046, 5.743634, 5.7364006, 5.747251, 5.7400174, 5.7906537, 5.732784, 5.671296, 5.7400174, 5.6640625, 5.6893806, 5.7038484, 5.656829, 5.7146993, 5.656829, 5.649595, 5.6640625, 5.642361, 5.649595, 5.711082, 5.6676793, 5.6893806, 5.6604457, 5.6315103, 5.642361, 5.6351275, 5.6532116, 5.5989585, 5.6387444, 5.5917244, 5.5989585, 5.5881076, 5.584491, 5.617043, 5.642361, 5.5664062, 5.570023, 5.5230036, 5.62066, 5.580874, 5.5555553, 5.584491, 5.5664062, 5.544705, 5.5374713, 5.5555553, 5.5266204, 5.5374713, 5.580874, 5.5157695, 5.5483217, 5.580874, 5.497685, 5.5013022, 5.497685, 5.5230036, 5.504919, 5.497685, 5.494068, 5.443432, 5.504919, 5.472367, 5.4615164, 5.472367, 5.4506655, 5.457899, 5.3855615, 5.3493924, 5.4144964, 5.4217305, 5.4217305, 5.403646, 5.396412, 5.3855615, 5.428964, 5.3855615, 5.4253473, 5.3819447, 5.3819447, 5.3240743, 5.36386, 5.3493924, 5.360243, 5.3855615, 5.353009, 5.3891783, 5.367477, 5.3747106, 5.3783274, 5.342159, 5.3023725, 5.3385415, 5.2625866, 5.266204, 5.31684, 5.320457, 5.3132234, 5.367477, 5.31684, 5.2372684, 5.295139, 5.2842884, 5.2734375, 5.251736, 5.2698207, 5.2698207, 5.2010994, 5.215567, 5.251736, 5.215567, -0.01808449, 2.0688658, 2.7307582, 3.3600984, 3.8519964, 3.9134839, 3.9026332, 3.8953993, 3.9171007, 3.9568865, 3.9568865, 3.9858217, 4.0039062, 4.018374, 3.9677372, 4.01114, 4.007523, 4.0509257, 4.021991, 4.079861, 4.184751, 4.181134, 4.094329, 4.1304975, 4.1413484, 4.191985, 4.1739006, 4.1775174, 4.170284, 4.2173033, 4.2064524, 4.271557, 4.2100697, 4.195602, 4.2896414, 4.271557, 4.32581, 4.307726, 4.300492, 4.296875, 4.333044, 4.401765, 4.3655963, 4.3511286, 4.3800635, 4.3945312, 4.445168, 4.434317, 4.37283, 4.5030384, 4.448785, 4.4524016, 4.5536747, 4.510272, 4.5645256, 4.546441, 4.575376, 4.575376, 4.5970774, 4.5645256, 4.5898438, 4.6296296, 4.622396, 4.658565, 4.6694155, 4.626013, 4.647714, 4.6694155, 4.7092013, 4.691117, 4.7417536, 4.7200522, 4.7345195, 4.814091, 4.8104744, 4.8828125, 4.799624, 4.8538775, 4.8719616, 4.824942, 4.9081306, 4.8936634, 4.951534, 4.9442997, 4.969618, 4.9840856, 4.9479165, 5.041956, 4.9985533, 5.027488, 5.00217, 5.1215277, 5.25897, 5.356626, 5.418113, 5.494068, 5.5989585, 5.6966147, 5.78342, 5.870226, 5.9895835, 6.047454, 6.188513, 6.275318, 6.3440394, 6.4850984, 6.600839, 6.6550927, 6.749132, 6.781684, 6.8757234, 7.0638022, 7.132523, 7.2265625, 7.2880497, 7.360388, 7.4797454, 7.559317, 7.66059, 7.7690973, 7.863137, 7.9716434, 8.083767, 8.1380205, 8.210359, 8.358651, 8.373119, 8.564815, 8.666088, 8.749276, 8.79268, 8.940972, 9.024161, 9.125434, 9.205006, 9.280961, 9.414786, 9.501592, 9.58478, 9.682436, 9.740307, 8.868634, 8.083767, 7.269965, 6.463397, 5.7689524, 5.8123555, 5.859375, 5.855758, 5.870226, 5.8919272, 5.8919272, 5.895544, 5.975116, 6.011285, 5.9570312, 6.0149016, 6.0040507, 6.072772, 6.076389, 6.069155, 6.0944734, 6.1306424, 6.199363, 6.1704283, 6.1631947, 6.184896, 6.199363, 6.213831, 6.2644677, 6.2717013, 6.3042536, 6.322338, 6.365741, 6.3440394, 6.3838253, 6.3802085, 6.4561634, 6.4091434, 6.4489293, 6.45978, 6.528501, 6.5067997, 6.532118, 6.528501, 6.589988, 6.5936055, 6.5719037, 6.5936055, 6.651476, 6.6731772, 6.702112, 6.712963, 6.7201967, 6.7093463, 6.828704, 6.7961516, 6.7853007, 6.8395543, 6.857639, 6.8974247, 6.8757234, 6.919126, 6.9516783, 6.9335938, 6.929977, 7.0167823, 7.0240164, 6.9733796, 7.056568, 7.042101, 7.168692, 7.146991, 7.1144385, 7.143374, 7.1650753, 7.1506076, 7.212095, 7.2157116, 7.2591147, 7.244647, 7.2916665, 7.309751, 7.2916665, 7.360388, 7.4001737, 7.3386865, 7.39294, 7.4146414, 7.4652777, 7.4544272, 7.483362, 7.494213, 7.4652777, 7.573785, 7.631655, 7.609954, 9.523293, 11.97555, 14.507379, 16.948784, 19.509548, 21.96904, 24.4864, 26.938658, 29.47772, 31.911892, 34.3967, 36.9647, 39.373554, 41.858364, 41.95602, 38.740597, 36.295574, 33.78183, 31.282553, 28.725405, 26.280382, 23.828125, 21.296297, 18.804253, 16.34838, 13.841869, 11.400463, 8.85055, 6.4489293, 5.9172454, 5.870226, 5.8521414, 5.794271, 5.7725697, 5.7761865, 5.7400174, 5.7291665, 5.707465, 5.6966147, 5.671296, 5.6676793, 5.642361, 5.617043, 5.6025753, 5.577257, 5.4868345, 5.5555553, 5.504919, 5.472367, 5.4506655, 5.439815, 5.3891783, 5.443432, 5.3493924, 5.342159, 5.360243, 5.3819447, 5.31684, 5.331308, 5.295139, 5.2842884, 5.2336516, 5.2336516, 5.1757812, 5.190249, 5.2119503, 5.1106772, 5.0962095, 5.067274, 5.10706, 5.0564237, 5.0600405, 4.9877024, 5.0094037, 4.962384, 4.966001, 4.962384, 4.9189816, 4.929832, 4.875579, 4.904514, 4.8430266, 4.8466434, 4.79239, 4.7743053, 4.7779226, 4.763455, 4.712818, 4.712818, 4.698351, 4.6730323, 4.6296296, 4.6694155, 4.636863, 4.5934606, 4.5572915, 4.5898438, 4.550058, 4.510272, 4.513889, 4.448785, 4.434317, 4.448785, 4.4162326, 4.3836803, 4.3438945, 4.412616, 4.3655963, 4.32581, 4.322193, 4.296875, 4.307726, 4.2643228, 4.2498555, 4.260706, 4.2136865, 4.184751, 4.148582, 4.1666665, 4.1739006, 4.0979457, 4.0509257, 4.1304975, 4.11603, 4.0400753, 4.05816, 4.043692, 3.9930556, 4.0002894, 3.9641204, 3.9134839, 3.9460359, 3.9315684, 3.8664641, 3.8809316, 3.8809316, 3.8628473, 3.870081, 3.765191, 3.8194444, 3.7760417, 3.761574, 3.7760417, 3.7145543, 3.7941263, 3.7217882, 3.768808, 3.7181714, 3.7109375, 3.685619, 3.653067, 3.6711516, 3.6747684, 3.6277487, 3.5951967, 3.653067, 3.5807292, 3.5771122, 3.5662615, 3.5879629, 3.5373263, 3.5264757, 3.4939237, 3.479456, 3.5083911, 3.4975405, 3.4541378, 3.4613714, 3.4288194, 3.446904, 3.3564816, 3.4288194, 3.414352, 3.3854167, 3.3926504, 3.3311632, 3.2769098, 3.3962674, 3.3275464, 3.305845, 3.3094618, 3.2443576, 3.2443576, 3.2913773, 3.200955, 3.1973379, 3.2118056, 3.193721, 3.200955, 3.1394675, 3.0960648, 3.1322339, 3.1286168, 3.0852141, 3.056279, 3.0635128, 3.0743635, 3.0635128, 3.0454283, 3.0092592, 3.0056424, 3.0092592, 2.9622395, 2.9658566, 2.980324, 2.9730902, 2.9333043, 2.9333043, 2.879051, 2.879051, 2.879051, 2.904369, 2.8284144, 2.81033, 2.7813947, 2.8211806, 2.8139467, 2.879051, 2.7596934, 2.7633102, 2.7271411, 2.7596934, 2.7090566, 2.6909723, 2.7235243, 2.6439526, 2.7162905, 2.633102, 2.6367188, 2.6439526, 2.6222513, 2.593316, 2.5499132, 2.6114004, 2.5860822, 2.5173612, 2.5752316, 2.4956598, 2.4920428, 2.5499132, 2.4920428, 2.4703414, 2.481192, 2.419705, 2.4414062, 2.44864, 2.3726852, 2.4016204, 2.419705, 2.34375, 2.4016204, 2.3654513, 2.34375, 2.3220487, 2.307581, 2.3148148, 2.3003473, 2.2967303, 2.2822628, 2.2243924, 2.199074, 1.9965278, 1.3599538, 0.77039933, 4.235388, 6.915509, 6.8323207, 6.8865743, 6.9082756, 6.922743, 6.919126, 6.9335938, 6.922743, 6.929977, 6.9082756, 6.9118924, 6.9372106, 6.966146, 6.9372106, 6.966146, 6.969763, 7.002315, 6.969763, 6.9733796, 6.922743, 6.9480615, 6.9516783, 6.9986978, 6.9625287, 6.966146, 7.0384836, 7.0167823, 7.0167823, 7.060185, 6.9769964, 7.027633, 7.020399, 7.042101, 7.034867, 7.107205, 7.0638022, 7.0529513, 6.995081, 7.0638022, 7.060185, 7.03125, 7.0891204, 7.1289062, 7.0891204, 7.0638022, 7.0638022, 7.042101, 7.056568, 7.1289062, 7.060185, 7.132523, 7.1144385, 7.1216726, 7.1216726, 7.1650753, 7.103588, 7.132523, 7.1252894, 7.1614585, 7.13614, 7.3423033, 7.9824944, 8.629919, 9.302662, 9.993489, 10.250289, 10.275608, 10.239439, 10.315393, 10.304543, 10.362413, 10.340712, 10.380498, 10.441985, 10.427517, 10.405816, 10.449219, 10.478154, 10.445601, 10.499855, 10.543258, 10.550492, 10.550492, 10.546875, 10.590278, 10.619213, 10.640914, 10.622829, 10.619213, 10.684318, 10.706018, 10.745805, 10.7421875, 10.821759, 10.771123, 10.767506, 10.774739, 10.821759, 10.8723955, 10.883246, 10.828993, 10.868779, 10.876013, 10.955585, 10.9375, 10.912182, 10.988136, 10.980903, 11.053241, 11.035156, 11.035156, 11.020689, 11.085793, 11.067708, 11.111111, 11.125579, 11.093026, 11.176215, 11.190682, 11.201533, 11.212384, 11.183449, 11.281105, 11.295573, 11.288339, 11.29919, 11.338976, 11.291956, 11.400463, 11.433015, 11.389612, 11.436632, 11.41493, 11.436632, 11.458333, 11.487268, 11.541522, 11.548756, 11.581307, 11.56684, 11.595776, 11.588542, 11.668114, 11.642796, 11.631945, 11.722367, 11.729601, 11.689815, 11.678964, 11.780237, 11.76577, 11.892361, 11.979167, 12.051505, 12.134693, 12.319155, 12.322772, 12.445746, 12.55787, 12.659143, 12.702546, 12.86169, 12.973814, 13.017217, 13.17636, 13.259548, 13.357204, 13.429543, 13.603154, 13.675492, 13.718895, 13.809318, 14.008246, 14.058883, 14.152923, 14.275897, 14.36632, 14.438658, 14.550781, 14.63397, 14.713542, 14.847367, 14.970342, 15.006511, 15.143952, 15.209057, 15.3464985, 15.476707, 15.5598955, 15.700954, 15.650318, 15.878182, 15.968605, 16.059029, 16.109665, 16.257957, 16.304977, 16.489439, 16.536459, 16.713686, 16.749855, 16.681135, 15.849248, 15.04268, 14.228877, 13.440393, 12.879774, 12.865307, 12.995515, 12.962963, 12.905092, 12.926794, 13.013599, 13.017217, 13.096788, 13.035301, 13.104022, 13.100405, 13.1691265, 13.190827, 13.17636, 13.179976, 13.212529, 13.205296, 13.230614, 13.263165, 13.255932, 13.284867, 13.306568, 13.357204, 13.353588, 13.317419, 13.418693, 13.422309, 13.451244, 13.494647, 13.49103, 13.5597515, 13.53805, 13.595921, 13.621239, 13.624855, 13.646557, 13.624855, 13.697193, 13.726129, 13.718895, 13.7369795, 13.762298, 13.798467, 13.751447, 13.838252, 13.812934, 13.86357, 13.903357, 13.870805, 13.986546, 13.972077, 13.935908, 14.019097, 14.044415, 14.0625, 14.1276045, 14.076967, 14.102286, 14.080585, 14.145689, 14.163774, 14.196325, 14.243345, 14.26143, 14.268663, 14.293982, 14.308449, 14.315682, 14.359086, 14.384404, 14.3880205, 14.637587, 17.12963, 19.545717, 22.106482, 24.594908, 27.02908, 29.542824, 32.00955, 34.49074, 37.01172, 39.50376, 41.923466, 41.927082, 38.925056, 36.342594, 33.778214, 31.369358, 28.884548, 26.425058, 23.969185, 21.45544, 18.927229, 16.536459, 14.026331, 12.742332, 12.666377, 12.641059, 12.684462, 12.572338, 12.579572, 12.594039, 12.514467, 12.478298, 12.471065, 12.521702, 12.416811, 12.413195, 12.3878765, 12.416811, 12.351707, 12.319155, 12.333623, 12.333623, 12.275752, 12.286603, 12.297454, 12.188947, 12.185329, 12.188947, 12.1744795, 12.185329, 12.160011, 12.073206, 12.112992, 12.069589, 12.069589, 11.968316, 12.037037, 11.942998, 11.924913, 11.903212, 11.877893, 11.895978, 11.885127, 11.877893, 11.798322, 11.780237, 11.736835, 11.77662, 11.736835, 11.682581, 11.668114, 11.689815, 11.646412, 11.6536455, 11.621094, 11.574074, 11.61386, 11.490886, 11.541522, 11.548756, 11.443866, 11.505353, 11.469184, 11.436632, 11.3932295, 11.371528, 11.3932295, 11.338976, 11.313658, 11.291956, 11.248553, 11.266638, 11.244936, 11.244936, 11.1943, 11.190682, 11.205151, 11.201533, 11.129195, 11.121962, 11.107494, 11.093026, 11.027923, 11.064092, 11.046007, 11.020689, 10.99537, 10.966435, 10.933883, 10.926649, 10.87963, 10.883246, 10.792824, 10.839844, 10.854311, 10.839844, 10.767506, 10.763889, 10.724103, 10.760272, 10.716869, 10.698785, 10.651765, 10.673467, 10.662616, 10.630064, 10.615596, 10.637298, 10.539641, 10.561342, 10.492621, 10.514323, 10.420283, 10.441985, 10.449219, 10.445601, 10.384114, 10.394965, 10.391349, 10.340712, 10.300926, 10.286458, 10.250289, 10.340712, 10.243055, 10.250289, 10.196036, 10.192419, 10.177952, 10.152633, 10.145399, 10.163484, 10.105614, 10.054976, 10.069445, 10.047743, 9.968171, 10.062211, 9.979022, 10.00434, 9.997107, 9.964555, 9.932002, 9.892217, 9.924768, 9.866899, 9.8307295, 9.812645, 9.765625, 9.743923, 9.780092, 9.751158, 9.74754, 9.704138, 9.628182, 9.689671, 9.660735, 9.613715, 9.635417, 9.620949, 9.559462, 9.516059, 9.544994, 9.606482, 9.483507, 9.505208, 9.447338, 9.490741, 9.4401045, 9.436487, 9.382234, 9.403935, 9.382234, 9.371383, 9.331597, 9.31713, 9.27011, 9.306279, 9.248408, 9.259259, 9.27011, 9.172454, 9.143518, 9.139901, 9.1796875, 9.129051, 9.089265, 9.078414, 9.092882, 9.078414, 9.01331, 9.0494795, 8.973524, 8.980758, 9.024161, 8.959057, 9.00246, 8.908421, 8.857783, 8.861401, 8.854167, 8.80353, 8.861401, 8.760127, 8.85055, 8.817998, 8.734809, 8.731193, 8.702257, 8.723958, 8.734809, 8.6588545, 8.619068, 8.615452, 8.608217, 8.579283, 8.503327, 7.8559027, 7.309751, 6.6333914, 5.964265, 5.530237, 5.541088, 5.5121527, 5.4759836, 5.533854, 5.5013022, 5.494068, 5.5013022, 5.5157695, 5.3855615, 5.4470487, 5.439815, 5.544705, 5.4615164, 5.443432, 5.360243, 5.4000287, 5.432581, 5.4000287, 5.367477, 5.4470487, 5.3710938, 5.4253473, 5.3783274, 5.396412, 5.4470487, 5.3240743, 5.3710938, 5.4108796, 5.4361978, 5.342159, 5.353009, 5.367477, 5.4000287, 5.392795, 5.4108796, 5.3059897, 5.331308, 5.3710938, 5.31684, 5.360243, 5.327691, 5.327691, 5.31684, 5.287905, 5.2228007, 5.3493924, 5.331308, 5.2987556, 5.255353, 5.3096066, 5.287905, 5.266204, 5.266204, 5.2119503, 5.2228007, 5.2408853, 5.2842884, 5.230035, 5.1974826, -0.047019675, 1.5661169, 5.5266204, 6.0583043, 6.0908566, 6.0583043, 6.141493, 6.1161747, 6.069155, 6.1631947, 6.076389, 6.101707, 6.141493, 6.1559606, 6.1595774, 6.112558, 6.1523438, 6.141493, 6.076389, 6.2065973, 6.1270256, 6.1053243, 6.101707, 6.1921296, 6.137876, 6.1812787, 6.137876, 6.174045, 6.1921296, 6.2282987, 6.260851, 6.174045, 6.260851, 6.174045, 6.2065973, 6.224682, 6.2427664, 6.246383, 6.2572336, 6.289786, 6.224682, 6.246383, 6.1812787, 6.2825522, 6.213831, 6.239149, 6.224682, 6.260851, 6.2680845, 6.2680845, 6.3042536, 6.253617, 6.2572336, 6.3295717, 6.246383, 6.3187213, 6.3404226, 6.3404226, 6.311487, 6.2717013, 6.325955, 6.286169, 6.278935, 6.87934, 7.494213, 8.11632, 8.828849, 9.371383, 9.414786, 9.461805, 9.505208, 9.483507, 9.461805, 9.566695, 9.476274, 9.566695, 9.592014, 9.58478, 9.642651, 9.58478, 9.689671, 9.711371, 9.671586, 9.67882, 9.646267, 9.696904, 9.74754, 9.790943, 9.787327, 9.812645, 9.85243, 9.841579, 9.863281, 9.866899, 9.89945, 9.884983, 9.950087, 9.953704, 9.997107, 9.979022, 9.993489, 10.047743, 10.0441265, 10.105614, 10.116464, 10.076678, 10.047743, 10.09838, 10.101996, 10.145399, 10.196036, 10.239439, 10.199653, 10.206886, 10.246673, 10.311776, 10.279224, 10.293693, 10.311776, 10.319011, 10.358796, 10.398582, 10.380498, 10.441985, 10.402199, 10.4817705, 10.409432, 10.478154, 10.445601, 10.590278, 10.507089, 10.590278, 10.536024, 10.56496, 10.583044, 10.648149, 10.608362, 10.695168, 10.6807, 10.698785, 10.771123, 10.716869, 10.807292, 10.756655, 10.818142, 10.8253765, 10.8723955, 10.814526, 10.915798, 10.886864, 10.962818, 10.933883, 10.9375, 11.024305, 11.08941, 11.168982, 11.273871, 11.422164, 11.487268, 11.577691, 11.66088, 11.791088, 11.942998, 12.004485, 12.051505, 12.116609, 12.2432, 12.380642, 12.449364, 12.597656, 12.680845, 12.764033, 12.847222, 12.948495, 13.064236, 13.147425, 13.245081, 13.378906, 13.418693, 13.610388, 13.646557, 13.70081, 13.8671875, 13.925057, 14.087818, 14.160156, 14.275897, 14.355469, 14.43504, 14.510995, 14.680989, 14.756945, 14.832899, 14.966724, 15.046296, 15.154803, 15.292245, 15.389901, 15.455006, 15.5598955, 15.628617, 15.794994, 15.867332, 15.954138, 15.353733, 14.612268, 13.7839985, 13.0027485, 12.123842, 12.076823, 12.087673, 12.094908, 12.09129, 12.120226, 12.203414, 12.178096, 12.160011, 12.203414, 12.250434, 12.268518, 12.311921, 12.3046875, 12.3046875, 12.340857, 12.337239, 12.380642, 12.398726, 12.416811, 12.481915, 12.492766, 12.528935, 12.460214, 12.525318, 12.518085, 12.561487, 12.550636, 12.572338, 12.644676, 12.662761, 12.69893, 12.706163, 12.720631, 12.70978, 12.745949, 12.771267, 12.767651, 12.843605, 12.8255205, 12.86169, 12.87254, 12.879774, 12.944879, 12.966579, 12.915943, 12.962963, 12.97743, 13.042535, 13.053386, 13.107639, 13.118489, 13.132957, 13.1691265, 13.12934, 13.198061, 13.194445, 13.248698, 13.263165, 13.274016, 13.292101, 13.321036, 13.342737, 13.3463545, 13.411458, 13.389757, 13.425926, 13.43316, 13.483796, 13.530816, 13.512732, 13.556134, 13.545283, 13.563368, 13.603154, 13.6067705, 13.697193, 13.671875, 13.715278, 13.722511, 13.733362, 13.762298, 13.827401, 13.776765, 13.859954, 13.870805, 13.899739, 13.914207, 13.91059, 13.943142, 13.91059, 14.001013, 14.9088545, 17.379196, 19.874855, 22.363281, 24.927662, 27.434172, 29.868345, 32.37124, 34.84158, 37.351707, 39.850983, 42.30324, 42.317707, 38.404224, 35.919415, 33.412907, 30.917246, 28.464989, 25.951244, 23.441116, 20.916521, 18.478733, 15.9505205, 13.469329, 11.038774, 10.152633, 10.141783, 10.0911455, 10.087529, 10.101996, 10.058594, 10.033276, 10.00434, 9.997107, 9.89945, 9.950087, 9.950087, 9.942853, 9.870515, 9.845197, 9.801794, 9.8307295, 9.798177, 9.790943, 9.790943, 9.725839, 9.664351, 9.7005205, 9.704138, 9.624566, 9.664351, 9.58478, 9.559462, 9.563079, 9.544994, 9.512443, 9.541377, 9.4871235, 9.454572, 9.425636, 9.447338, 9.396702, 9.382234, 9.360533, 9.346065, 9.342448, 9.331597, 9.3098955, 9.288195, 9.212239, 9.241175, 9.172454, 9.215857, 9.168837, 9.154369, 9.132668, 9.092882, 9.027778, 9.092882, 9.024161, 8.984375, 8.987992, 8.948206, 8.908421, 8.937355, 8.875868, 8.893952, 8.861401, 8.854167, 8.828849, 8.832465, 8.817998, 8.756511, 8.785445, 8.770978, 8.709491, 8.655237, 8.74566, 8.6588545, 8.648004, 8.626302, 8.644386, 8.579283, 8.586516, 8.485243, 8.532263, 8.452691, 8.5286455, 8.492476, 8.445457, 8.39482, 8.420139, 8.387587, 8.39482, 8.351418, 8.347801, 8.318866, 8.326099, 8.224827, 8.260995, 8.217592, 8.188658, 8.192274, 8.217592, 8.098235, 8.083767, 8.0910015, 8.065682, 8.065682, 8.051215, 8.051215, 8.076533, 8.015046, 7.9716434, 7.953559, 7.9354744, 7.91739, 7.913773, 7.913773, 7.884838, 7.808883, 7.787182, 7.7907987, 7.8197336, 7.8197336, 7.761863, 7.7582464, 7.700376, 7.7148438, 7.6822915, 7.685909, 7.6461225, 7.6208043, 7.570168, 7.5882525, 7.5882525, 7.5050635, 7.562934, 7.533999, 7.526765, 7.4688945, 7.472512, 7.49783, 7.421875, 7.425492, 7.349537, 7.4037905, 7.3531537, 7.3748555, 7.306134, 7.3314524, 7.3025174, 7.313368, 7.2012444, 7.2229457, 7.295284, 7.248264, 7.172309, 7.172309, 7.1614585, 7.13614, 7.0855036, 7.0746527, 7.0891204, 7.0493345, 7.071036, 7.0167823, 6.966146, 6.9516783, 6.9516783, 6.9118924, 6.922743, 6.8684897, 6.8757234, 6.8250866, 6.8757234, 6.8684897, 6.8033853, 6.7997684, 6.781684, 6.6876445, 6.756366, 6.6948786, 6.6948786, 6.7274303, 6.6731772, 6.680411, 6.6587095, 6.6225405, 6.5863714, 6.604456, 6.575521, 6.5863714, 6.5538197, 6.5212674, 6.4742475, 6.499566, 6.4489293, 6.4344616, 6.4814816, 6.35489, 6.358507, 6.362124, 6.3368053, 6.311487, 6.358507, 6.2717013, 6.289786, 6.2572336, 6.224682, 6.213831, 6.2355323, 6.184896, 6.184896, 6.1812787, 6.09809, 6.1161747, 6.137876, 6.112558, 6.0872397, 6.0257525, 6.0293694, 6.032986, 6.101707, 5.964265, 5.9787326, 5.9497976, 5.964265, 5.910012, 5.910012, 5.862992, 5.9172454, 5.834057, 5.8268228, 5.754485, 5.8376737, 5.787037, 5.7255497, 5.0311055, 4.4958043, 3.8664641, 3.1539352, 2.6511862, 2.6692708, 2.6475694, 2.6692708, 2.7379918, 2.6620371, 2.6837385, 2.6692708, 2.6692708, 2.6114004, 2.6367188, 2.6620371, 2.5788484, 2.6367188, 2.6186342, 2.6150174, 2.6077836, 2.6077836, 2.596933, 2.589699, 2.557147, 2.589699, 2.629485, 2.5788484, 2.6041667, 2.6186342, 2.5499132, 2.5607638, 2.5282118, 2.5354457, 2.589699, 2.6041667, 2.524595, 2.5028934, 2.4739583, 2.4956598, 2.513744, 2.524595, 2.5028934, 2.524595, 2.5065105, 2.5028934, 2.513744, 2.4594908, 2.4594908, 2.419705, 2.4739583, 2.5282118, 2.4414062, 2.4269388, 2.5028934, 2.4377894, 2.4594908, 2.4414062, 2.3943865, 2.4631076, 2.5028934, 2.445023, 2.4305556, 2.4377894, 0.0];
END_VAR
